// TIA Portal V20 export
// export: Created 2026-10-20T18:55:54.5785311Z, ExportSetting None, DisplayName Totally Integrated Automation Portal, DisplayVersion V20 Update 6, DisplayName TIA Portal Openness, DisplayVersion V20 Update 6, DisplayName TIA Portal Version Control Interface, DisplayVersion V20 Update 6, DisplayName SINAMICS Startdrive Advanced, DisplayVersion V20 SP1, DisplayName SINAMICS Startdrive G130, G150, S120, S150, SINAMICS MV, G220, S200, S210, DisplayVersion V20 SP1, DisplayName SINAMICS Startdrive G110M, G120, G120C, G120D, G120P, G115D, DisplayVersion V20 SP1, DisplayName STEP 7 Professional, DisplayVersion V20 Update 6, DisplayName STEP 7 Safety, DisplayVersion V20 Update 2, DisplayName WinCC Basic/Comfort/Advanced, DisplayVersion V20 Update 6, DisplayName WinCC Unified, DisplayVersion V20 Update 6
VAR_GLOBAL   // PLC tag table "Lock_8"
   Lock_8_Closed_CH1 AT %I1814.0 : Bool;
   Lock_8_Estop_CH1 AT %I1814.2 : Bool;
   "Lock Reset_8" AT %Q1496.0 : Bool;
   Lamps_8 AT %QB1494 : Byte;
   Lock_8_Closed_CH2 AT %I1814.1 : Bool;
   Lock_8_Estop_CH2 AT %I1814.3 : Bool;
   "Solenoid Enable_8" AT %Q1495.0 : Bool;
   Switches_8 AT %IB1346 : Byte;
   Lock_8_Reset_Input1 AT %Q1815.0 : Bool;
   Lock_8_Reset_Input3 AT %Q1815.2 : Bool;
   Lock_8_Reset_Input4 AT %Q1815.3 : Bool;
   Lock_8_Reset_Input2 AT %Q1815.1 : Bool;
   "Lock Position_8" AT %I1495.0 : Bool;
   "Guard Position_8" AT %I1494.0 : Bool;
END_VAR
